Universal Robots URScript: T005_deepseek-coder-v2_16b-lite-instruct-q4_K_M_baseline_rep2.urscript

# Define the home position
def home_position():
    movej([0.0, -1.5708, 1.5708, -1.5708, 1.5708, 0.0], 150.0, 0.5, 0)

# Define the approach position
def approach_position():
    movej([0.0, -1.5708, 1.5708, -1.5708, 1.5708, 0.0], 130.0, 0.5, 0)

# Define the descent position
def descent_position():
    movej([0.0, -1.5708, 1.5708, -1.5708, 1.5708, 0.0], 80.0, 0.5, 0)

# Define the scan line 1 position
def scan_line_1():
    movel([0.0, -0.2, 0.0, 0.0, 0.0, 0.0], [0.0, 0.0, -0.1, 0.0, 0.0, 0.0], 50.0, 0.5, 0)

# Define the scan line 2 position
def scan_line_2():
    movel([0.0, 0.2, 0.0, 0.0, 0.0, 0.0], [0.0, 0.0, -0.1, 0.0, 0.0, 0.0], 80.0, 0.5, 0)

# Define the scan line 3 position
def scan_line_3():
    movel([0.0, 0.2, 0.0, 0.0, 0.0, 0.0], [0.0, 0.0, -0.1, 0.0, 0.0, 0.0], 50.0, 0.5, 0)

# Define the scan line 4 position
def scan_line_4():
    movel([0.0, -0.2, 0.0, 0.0, 0.0, 0.0], [0.0, 0.0, -0.1, 0.0, 0.0, 0.0], 80.0, 0.5, 0)

# Define the scan line 5 position
def scan_line_5():
    movel([0.0, -0.2, 0.0, 0.0, 0.0, 0.0], [0.0, 0.0, -0.1, 0.0, 0.0, 0.0], 50.0, 0.5, 0)

# Main program
home_position()
approach_position()
descent_position()
scan_line_1()
scan_line_2()
scan_line_3()
scan_line_4()
scan_line_5()
